{attribute 'pack_mode' := '1'}
TYPE ST_PcsConfigWirePacket :
STRUCT
	Header	:	ST_MqttCommandHeader;
	Records	:	ARRAY[0..GVL_PARAM.PCS_COUNT-1] OF ST_PcsConfig_Rx;
END_STRUCT
END_TYPE

(* stored: Version 1.1.0.1, ProductVersion 3.1.4024.15
   DUT ST_PcsConfigWirePacket: Id {8618be98-f928-4405-88d3-f6ceeceaf96e} *)
